(* IEC 61131-3 sources: rusty/tests/lit/single/expressions, 5 files *)

(* ---- unsigned_comparison.st ---- *)
// RUN: %COMPILE %s && %RUN | %CHECK %s
//
// Two unsigned operands compare as unsigned values, also when a value has the highest bit set and
// no wider type is involved: UDINT with UDINT, and ULINT with ULINT or with a positive literal.

FUNCTION main
    VAR
        small_udint : UDINT := 5;
        large_udint : UDINT := 16#8000_0000;
        small_ulint : ULINT := 5;
        large_ulint : ULINT := 16#8000_0000_0000_0000;
    END_VAR
    printf('udint <: %d$N', small_udint < large_udint);
    printf('udint >: %d$N', large_udint > small_udint);
    printf('udint <=: %d$N', large_udint <= small_udint);
    printf('udint >=: %d$N', large_udint >= small_udint);
    // CHECK:      udint <: 1
    // CHECK-NEXT: udint >: 1
    // CHECK-NEXT: udint <=: 0
    // CHECK-NEXT: udint >=: 1

    printf('ulint <: %d$N', small_ulint < large_ulint);
    printf('ulint >: %d$N', large_ulint > small_ulint);
    printf('ulint <=: %d$N', large_ulint <= small_ulint);
    printf('ulint >=: %d$N', large_ulint >= small_ulint);
    // CHECK-NEXT: ulint <: 1
    // CHECK-NEXT: ulint >: 1
    // CHECK-NEXT: ulint <=: 0
    // CHECK-NEXT: ulint >=: 1

    printf('ulint > 5: %d$N', large_ulint > 5);
    // CHECK-NEXT: ulint > 5: 1
END_FUNCTION

(* ---- unsigned_comparison_bit_strings.st ---- *)
// RUN: %COMPILE %s && %RUN | %CHECK %s
//
// Two bit strings of the same type compare as unsigned values, also when a value has the highest
// bit set.

FUNCTION main
    VAR
        byte_low : BYTE := 1;
        byte_high : BYTE := 16#FF;
        word_low : WORD := 1;
        word_high : WORD := 16#FFFF;
        dword_low : DWORD := 1;
        dword_high : DWORD := 16#FFFF_FFFF;
        lword_low : LWORD := 1;
        lword_high : LWORD := 16#FFFF_FFFF_FFFF_FFFF;
    END_VAR
    printf('byte: %d$N', byte_high > byte_low);
    printf('word: %d$N', word_high > word_low);
    printf('dword: %d$N', dword_high > dword_low);
    printf('lword: %d$N', lword_high > lword_low);
    // CHECK:      byte: 1
    // CHECK-NEXT: word: 1
    // CHECK-NEXT: dword: 1
    // CHECK-NEXT: lword: 1
END_FUNCTION

(* ---- unsigned_comparison_multiple_operands.st ---- *)
// RUN: %COMPILE %s && %RUN | %CHECK %s
//
// Expressions with three and four operands compare an unsigned operand of 32 bits as an unsigned
// value in every comparison, with literals and with other unsigned operands.

FUNCTION main
    VAR
        a : UDINT := 16#8000_0000;
        b : UDINT := 5;
        c : UDINT := 1;
        d : UDINT := 0;
    END_VAR
    printf('a > 1 AND a < 16#FFFF_FFFF: %d$N', a > 1 AND a < 16#FFFF_FFFF);
    printf('a > b AND b > c AND c > d: %d$N', a > b AND b > c AND c > d);
    printf('a >= 16#8000_0000 OR a < 5: %d$N', a >= 16#8000_0000 OR a < 5);
    printf('((a > b) < c) > d: %d$N', ((a > b) < c) > d);
    printf('((a > b) = (b < a)) > d: %d$N', ((a > b) = (b < a)) > d);
    // CHECK:      a > 1 AND a < 16#FFFF_FFFF: 1
    // CHECK-NEXT: a > b AND b > c AND c > d: 1
    // CHECK-NEXT: a >= 16#8000_0000 OR a < 5: 1
    // CHECK-NEXT: ((a > b) < c) > d: 0
    // CHECK-NEXT: ((a > b) = (b < a)) > d: 1
END_FUNCTION

(* ---- unsigned_comparison_with_literal.st ---- *)
// RUN: %COMPILE %s && %RUN | %CHECK %s
//
// An unsigned operand of 32 or 64 bits compares with an integer literal as an unsigned value, also
// when the operand has the highest bit set.

FUNCTION main
    VAR
        udint_high : UDINT := 16#8000_0000;
        dword_high : DWORD := 16#8000_0000;
        ulint_high : ULINT := 16#8000_0000_0000_0000;
        lword_high : LWORD := 16#8000_0000_0000_0000;
    END_VAR
    printf('udint > 5: %d$N', udint_high > 5);
    printf('udint < 5: %d$N', udint_high < 5);
    printf('dword > 16#7FFF_FFFF: %d$N', dword_high > 16#7FFF_FFFF);
    printf('ulint > 5: %d$N', ulint_high > 5);
    printf('lword > 5: %d$N', lword_high > 5);
    // CHECK:      udint > 5: 1
    // CHECK-NEXT: udint < 5: 0
    // CHECK-NEXT: dword > 16#7FFF_FFFF: 1
    // CHECK-NEXT: ulint > 5: 1
    // CHECK-NEXT: lword > 5: 1
END_FUNCTION

(* ---- unary_plus.st ---- *)
// RUN: %COMPILE %s && %RUN | %CHECK %s

VAR_GLOBAL CONSTANT g1 : INT := +5; END_VAR

PROGRAM prog
VAR
    x : INT := +g1;
END_VAR
    // CHECK: 5
    printf('%d$N', x);
    +x;
    x := +x + 4;
    // CHECK: 9
    printf('%d$N', x);
    x := +-4 + 5;
    // CHECK: 1
    printf('%d$N', x);
    +-x;
    x := +foo(+x);
    // CHECK: 3
    printf('%d$N', x);
END_PROGRAM

FUNCTION foo : INT
VAR_INPUT
    x : INT;
END_VAR
    foo := +x + +2 - +(+x - +1);
END_FUNCTION

FUNCTION main
    prog();
END_FUNCTION
